(* IEC 61131-3 sources: kns-port-domestic/upstream/kns-pump-station/src/POUs/Log/F_EventCsvLine, 2 files *)

(* ---- F_EventCsvLine.decl.st ---- *)
// Назначение: строка CSV журнала (ASCII, «;», CRLF): seq;time_utc;kind;id;code;priority;old_state;new_state;
//             reason;value — номер, UTC ISO 8601 (пусто без часов), alarm/station, номер, код F_AlarmCode,
//             числовые значения перечислений, значение REAL_TO_STRING. Русский текст подставляет
//             tools_project/eventlog_decode.py на хосте.
// Автор:      kr0nsch
// Версия:     0.1.0
// Документ:   docs/DESIGN.md, раздел 9.2
FUNCTION F_EventCsvLine : STRING(GVL_Const.LOG_CSV_LINE_LEN)
VAR_INPUT
    stRecord : ST_EventRecord;      // запись журнала
END_VAR
VAR
    sKind : STRING(GVL_Const.LOG_SUFFIX_LEN);   // вид записи
    sHead : STRING(GVL_Const.LOG_CSV_LINE_LEN); // seq;time_utc;kind;id;code;
    sTail : STRING(GVL_Const.LOG_CSV_LINE_LEN); // priority;old_state;new_state;reason;
END_VAR
VAR CONSTANT
    SEP  : STRING := ';';
    CRLF : STRING := '$R$N';
END_VAR

(* ---- F_EventCsvLine.impl.st ---- *)
IF stRecord.eKind = E_EventKind.Alarm THEN
    sKind := 'alarm';
ELSE
    sKind := 'station';
END_IF
// seq;time_utc;kind;id;code;
sHead := CONCAT(CONCAT(UDINT_TO_STRING(stRecord.udiSeq), SEP),
                CONCAT(F_UtcToIso(uliUtc_ms := stRecord.uliUtc_ms), SEP));
sHead := CONCAT(sHead, CONCAT(CONCAT(sKind, SEP), CONCAT(UDINT_TO_STRING(stRecord.udiId), SEP)));
sHead := CONCAT(sHead, CONCAT(F_AlarmCode(udiId := stRecord.udiId), SEP));
// priority;old_state;new_state;reason;value
sTail := CONCAT(CONCAT(INT_TO_STRING(TO_INT(stRecord.ePriority)), SEP),
                CONCAT(INT_TO_STRING(TO_INT(stRecord.eOldState)), SEP));
sTail := CONCAT(sTail, CONCAT(CONCAT(INT_TO_STRING(TO_INT(stRecord.eNewState)), SEP),
                              CONCAT(INT_TO_STRING(TO_INT(stRecord.eReason)), SEP)));
F_EventCsvLine := CONCAT(CONCAT(sHead, sTail), CONCAT(REAL_TO_STRING(stRecord.rValue), CRLF));
